// Mitsubishi GX Works2 project: V2   PLC: FX3U/FX3UC

PROGRAM MAIN
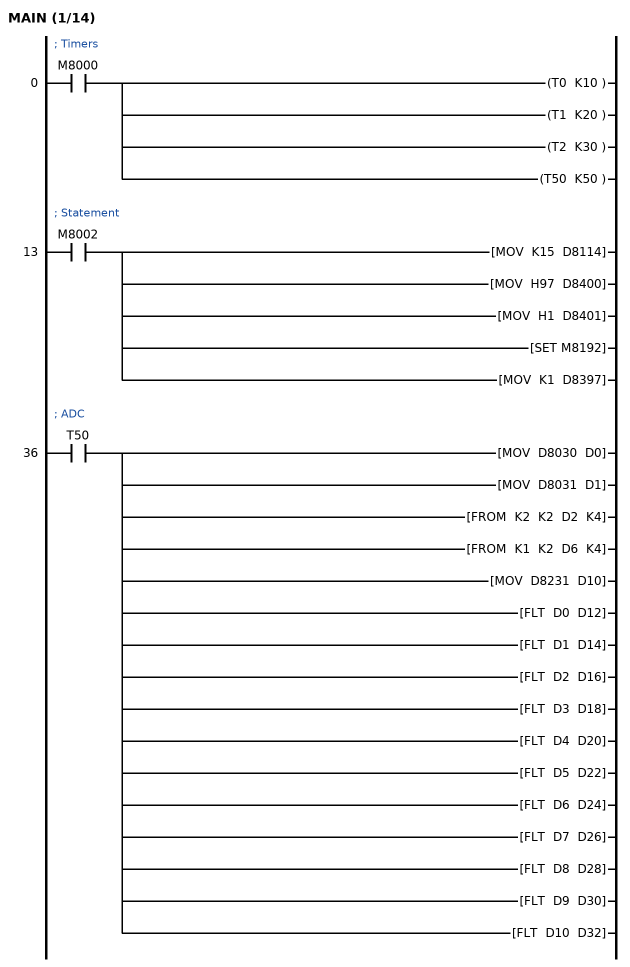
; Timers
0     LD      M8000
      OUT     T0 K10
      OUT     T1 K20
      OUT     T2 K30
      OUT     T50 K50
; Statement
13    LD      M8002
      MOV     K15 D8114
      MOV     H97 D8400
      MOV     H1 D8401
      SET     M8192
      MOV     K1 D8397
; ADC
36    LD      T50
      MOV     D8030 D0
      MOV     D8031 D1
      FROM    K2 K2 D2 K4
      FROM    K1 K2 D6 K4
      MOV     D8231 D10
      FLT     D0 D12
      FLT     D1 D14
      FLT     D2 D16
      FLT     D3 D18
      FLT     D4 D20
      FLT     D5 D22
      FLT     D6 D24
      FLT     D7 D26
      FLT     D8 D28
      FLT     D9 D30
      FLT     D10 D32
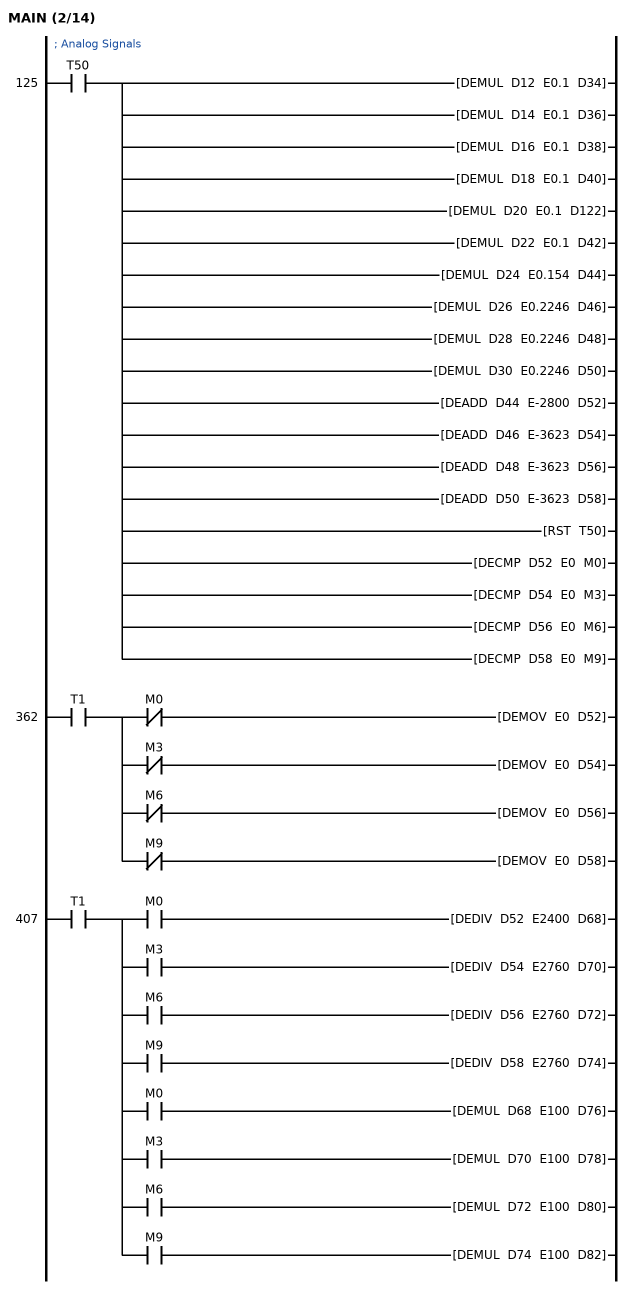
; Analog Signals
125   LD      T50
      DEMUL   D12 E0.1 D34
      DEMUL   D14 E0.1 D36
      DEMUL   D16 E0.1 D38
      DEMUL   D18 E0.1 D40
      DEMUL   D20 E0.1 D122
      DEMUL   D22 E0.1 D42
      DEMUL   D24 E0.154 D44
      DEMUL   D26 E0.2246 D46
      DEMUL   D28 E0.2246 D48
      DEMUL   D30 E0.2246 D50
      DEADD   D44 E-2800 D52
      DEADD   D46 E-3623 D54
      DEADD   D48 E-3623 D56
      DEADD   D50 E-3623 D58
      RST     T50
      DECMP   D52 E0 M0
      DECMP   D54 E0 M3
      DECMP   D56 E0 M6
      DECMP   D58 E0 M9
362   LD      T1
      MPS
      ANI     M0
      DEMOV   E0 D52
      MRD
      ANI     M3
      DEMOV   E0 D54
      MRD
      ANI     M6
      DEMOV   E0 D56
      MPP
      ANI     M9
      DEMOV   E0 D58
407   LD      T1
      MPS
      AND     M0
      DEDIV   D52 E2400 D68
      MRD
      AND     M3
      DEDIV   D54 E2760 D70
      MRD
      AND     M6
      DEDIV   D56 E2760 D72
      MRD
      AND     M9
      DEDIV   D58 E2760 D74
      MRD
      AND     M0
      DEMUL   D68 E100 D76
      MRD
      AND     M3
      DEMUL   D70 E100 D78
      MRD
      AND     M6
      DEMUL   D72 E100 D80
      MPP
      AND     M9
      DEMUL   D74 E100 D82
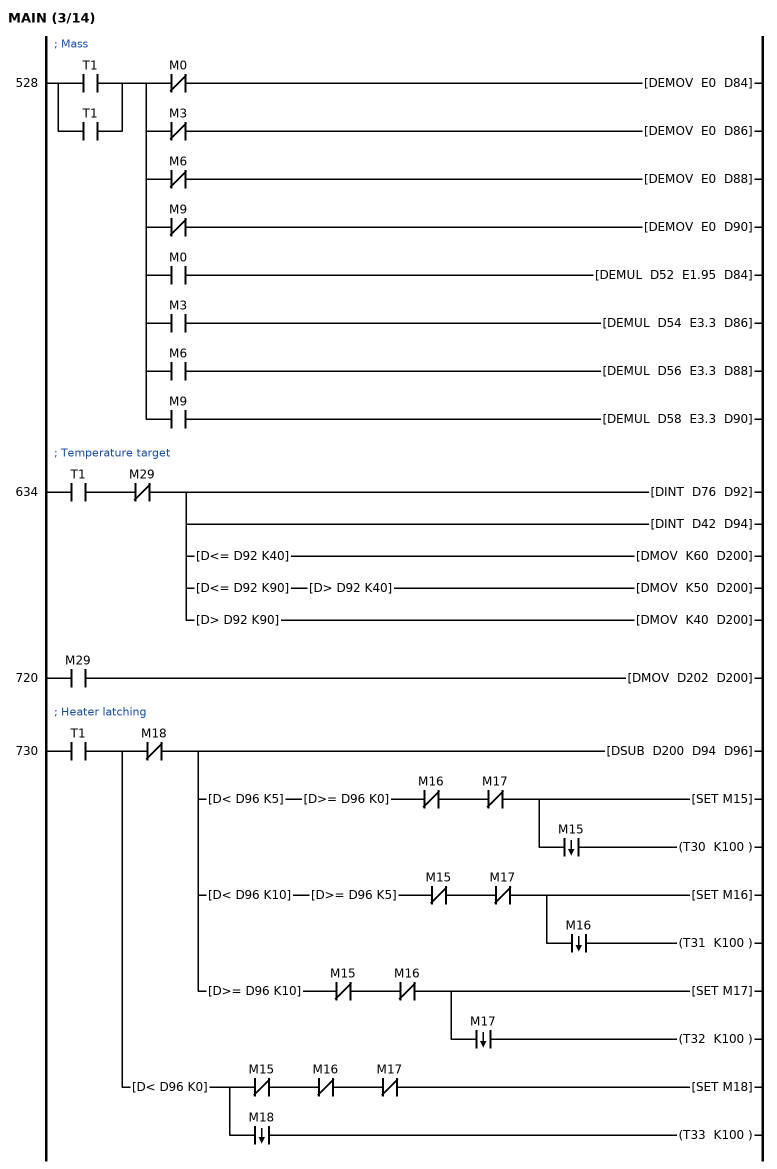
; Mass
528   LD      T1
      OR      T1
      MPS
      ANI     M0
      DEMOV   E0 D84
      MRD
      ANI     M3
      DEMOV   E0 D86
      MRD
      ANI     M6
      DEMOV   E0 D88
      MRD
      ANI     M9
      DEMOV   E0 D90
      MRD
      AND     M0
      DEMUL   D52 E1.95 D84
      MRD
      AND     M3
      DEMUL   D54 E3.3 D86
      MRD
      AND     M6
      DEMUL   D56 E3.3 D88
      MPP
      AND     M9
      DEMUL   D58 E3.3 D90
; Temperature target
634   LD      T1
      ANI     M29
      DINT    D76 D92
      DINT    D42 D94
      MPS
      ANDD<=  D92 K40
      DMOV    K60 D200
      MRD
      ANDD<=  D92 K90
      ANDD>   D92 K40
      DMOV    K50 D200
      MPP
      ANDD>   D92 K90
      DMOV    K40 D200
720   LD      M29
      DMOV    D202 D200
; Heater latching
730   LD      T1
      MPS
      ANI     M18
      DSUB    D200 D94 D96
      MPS
      ANDD<   D96 K5
      ANDD>=  D96 K0
      ANI     M16
      ANI     M17
      SET     M15
      ANDF    M15
      OUT     T30 K100
      MRD
      ANDD<   D96 K10
      ANDD>=  D96 K5
      ANI     M15
      ANI     M17
      SET     M16
      ANDF    M16
      OUT     T31 K100
      MPP
      ANDD>=  D96 K10
      ANI     M15
      ANI     M16
      SET     M17
      ANDF    M17
      OUT     T32 K100
      MPP
      ANDD<   D96 K0
      MPS
      ANI     M15
      ANI     M16
      ANI     M17
      SET     M18
      MPP
      ANDF    M18
      OUT     T33 K100
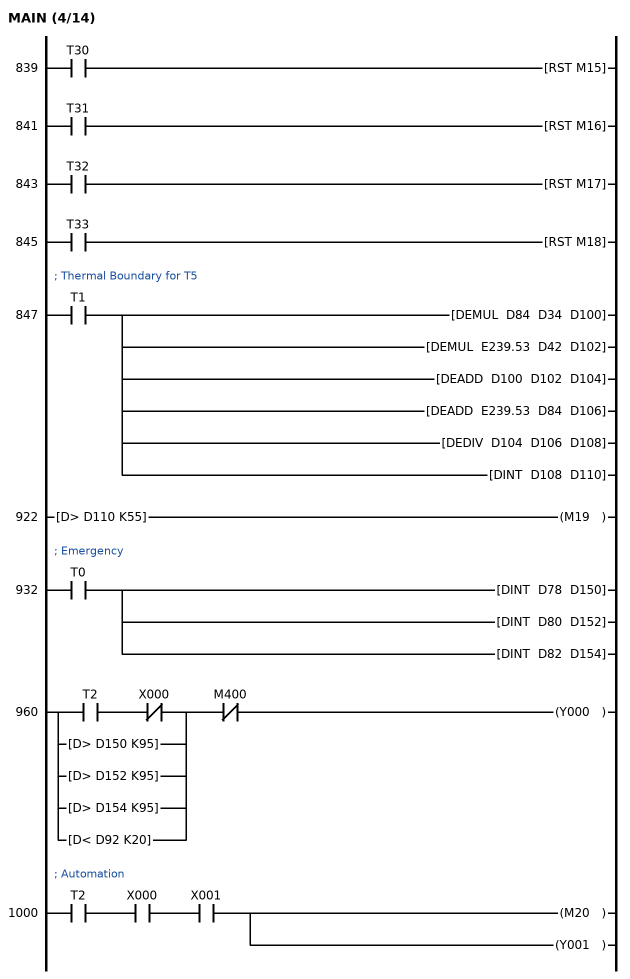
839   LD      T30
      RST     M15
841   LD      T31
      RST     M16
843   LD      T32
      RST     M17
845   LD      T33
      RST     M18
; Thermal Boundary for T5
847   LD      T1
      DEMUL   D84 D34 D100
      DEMUL   E239.53 D42 D102
      DEADD   D100 D102 D104
      DEADD   E239.53 D84 D106
      DEDIV   D104 D106 D108
      DINT    D108 D110
922   LDD>    D110 K55
      OUT     M19
; Emergency
932   LD      T0
      DINT    D78 D150
      DINT    D80 D152
      DINT    D82 D154
960   LD      T2
      ANI     X000
      ORD>    D150 K95
      ORD>    D152 K95
      ORD>    D154 K95
      ORD<    D92 K20
      ANI     M400
      OUT     Y000
; Automation
1000  LD      T2
      AND     X000
      AND     X001
      OUT     M20
      OUT     Y001
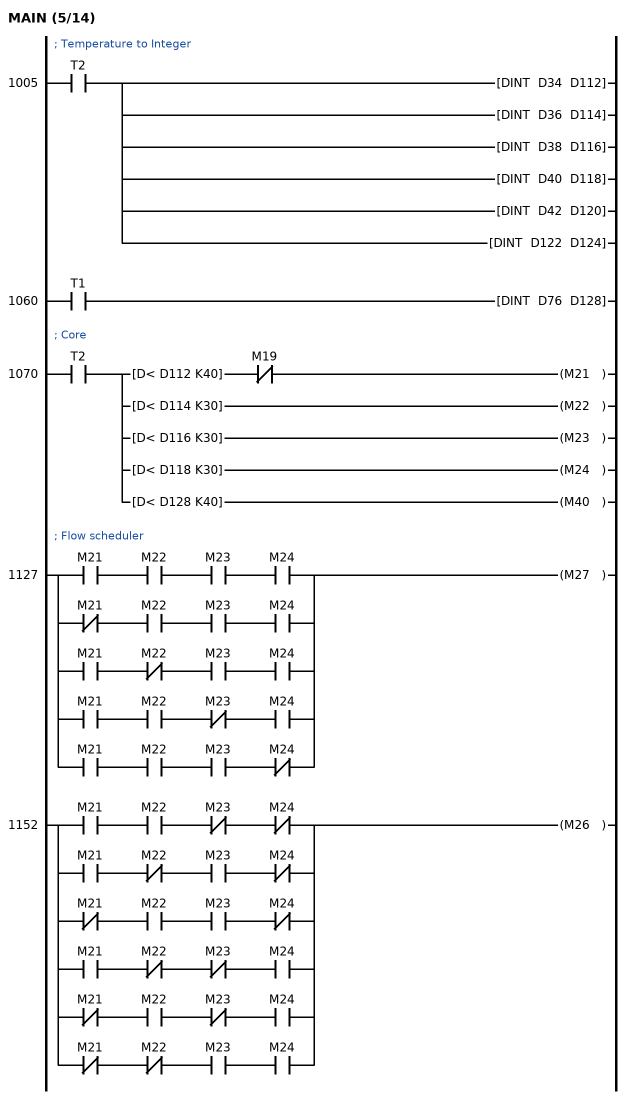
; Temperature to Integer
1005  LD      T2
      DINT    D34 D112
      DINT    D36 D114
      DINT    D38 D116
      DINT    D40 D118
      DINT    D42 D120
      DINT    D122 D124
1060  LD      T1
      DINT    D76 D128
; Core
1070  LD      T2
      MPS
      ANDD<   D112 K40
      ANI     M19
      OUT     M21
      MRD
      ANDD<   D114 K30
      OUT     M22
      MRD
      ANDD<   D116 K30
      OUT     M23
      MRD
      ANDD<   D118 K30
      OUT     M24
      MPP
      ANDD<   D128 K40
      OUT     M40
; Flow scheduler
1127  LD      M21
      AND     M22
      AND     M23
      AND     M24
      LDI     M21
      AND     M22
      AND     M23
      AND     M24
      ORB
      LD      M21
      ANI     M22
      AND     M23
      AND     M24
      ORB
      LD      M21
      AND     M22
      ANI     M23
      AND     M24
      ORB
      LD      M21
      AND     M22
      AND     M23
      ANI     M24
      ORB
      OUT     M27
1152  LD      M21
      AND     M22
      ANI     M23
      ANI     M24
      LD      M21
      ANI     M22
      AND     M23
      ANI     M24
      ORB
      LDI     M21
      AND     M22
      AND     M23
      ANI     M24
      ORB
      LD      M21
      ANI     M22
      ANI     M23
      AND     M24
      ORB
      LDI     M21
      AND     M22
      ANI     M23
      AND     M24
      ORB
      LDI     M21
      ANI     M22
      AND     M23
      AND     M24
      ORB
      OUT     M26
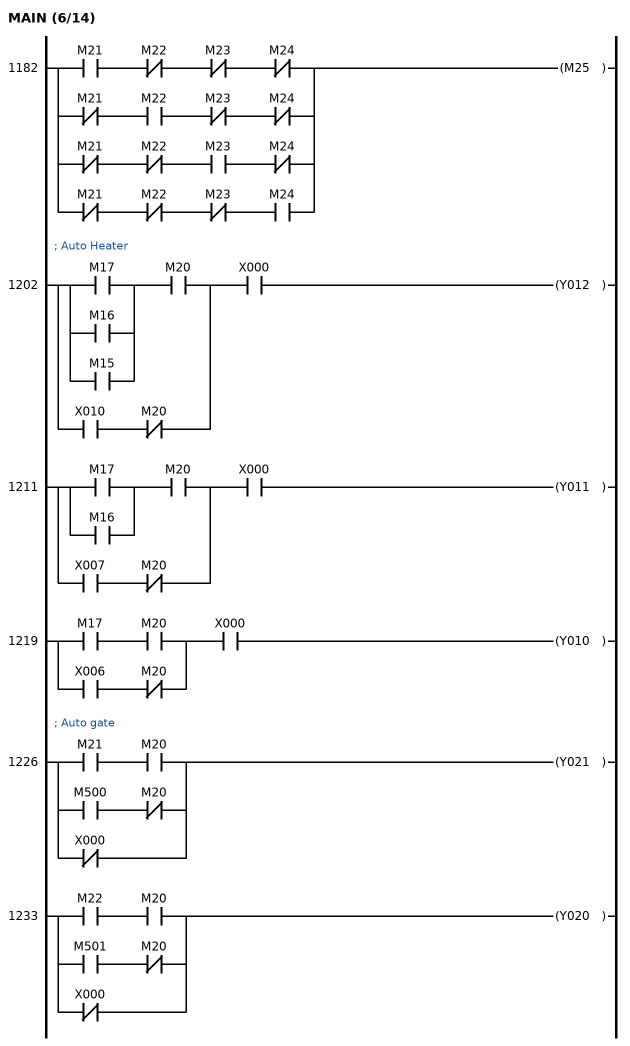
1182  LD      M21
      ANI     M22
      ANI     M23
      ANI     M24
      LDI     M21
      AND     M22
      ANI     M23
      ANI     M24
      ORB
      LDI     M21
      ANI     M22
      AND     M23
      ANI     M24
      ORB
      LDI     M21
      ANI     M22
      ANI     M23
      AND     M24
      ORB
      OUT     M25
; Auto Heater
1202  LD      M17
      OR      M16
      OR      M15
      AND     M20
      LD      X010
      ANI     M20
      ORB
      AND     X000
      OUT     Y012
1211  LD      M17
      OR      M16
      AND     M20
      LD      X007
      ANI     M20
      ORB
      AND     X000
      OUT     Y011
1219  LD      M17
      AND     M20
      LD      X006
      ANI     M20
      ORB
      AND     X000
      OUT     Y010
; Auto gate
1226  LD      M21
      AND     M20
      LD      M500
      ANI     M20
      ORB
      ORI     X000
      OUT     Y021
1233  LD      M22
      AND     M20
      LD      M501
      ANI     M20
      ORB
      ORI     X000
      OUT     Y020
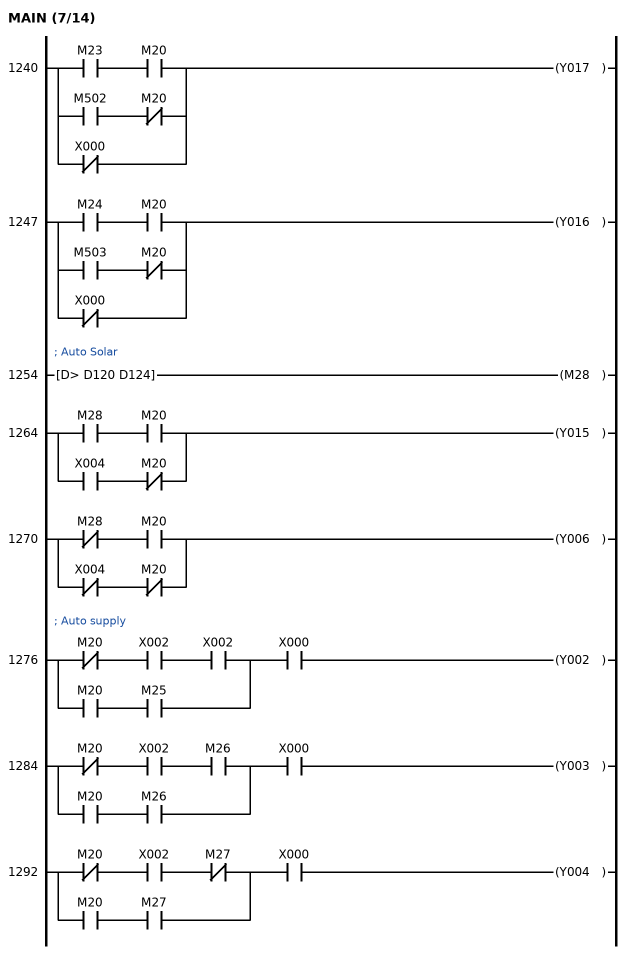
1240  LD      M23
      AND     M20
      LD      M502
      ANI     M20
      ORB
      ORI     X000
      OUT     Y017
1247  LD      M24
      AND     M20
      LD      M503
      ANI     M20
      ORB
      ORI     X000
      OUT     Y016
; Auto Solar
1254  LDD>    D120 D124
      OUT     M28
1264  LD      M28
      AND     M20
      LD      X004
      ANI     M20
      ORB
      OUT     Y015
1270  LDI     M28
      AND     M20
      LDI     X004
      ANI     M20
      ORB
      OUT     Y006
; Auto supply
1276  LDI     M20
      AND     X002
      AND     X002
      LD      M20
      AND     M25
      ORB
      AND     X000
      OUT     Y002
1284  LDI     M20
      AND     X002
      AND     M26
      LD      M20
      AND     M26
      ORB
      AND     X000
      OUT     Y003
1292  LDI     M20
      AND     X002
      ANI     M27
      LD      M20
      AND     M27
      ORB
      AND     X000
      OUT     Y004
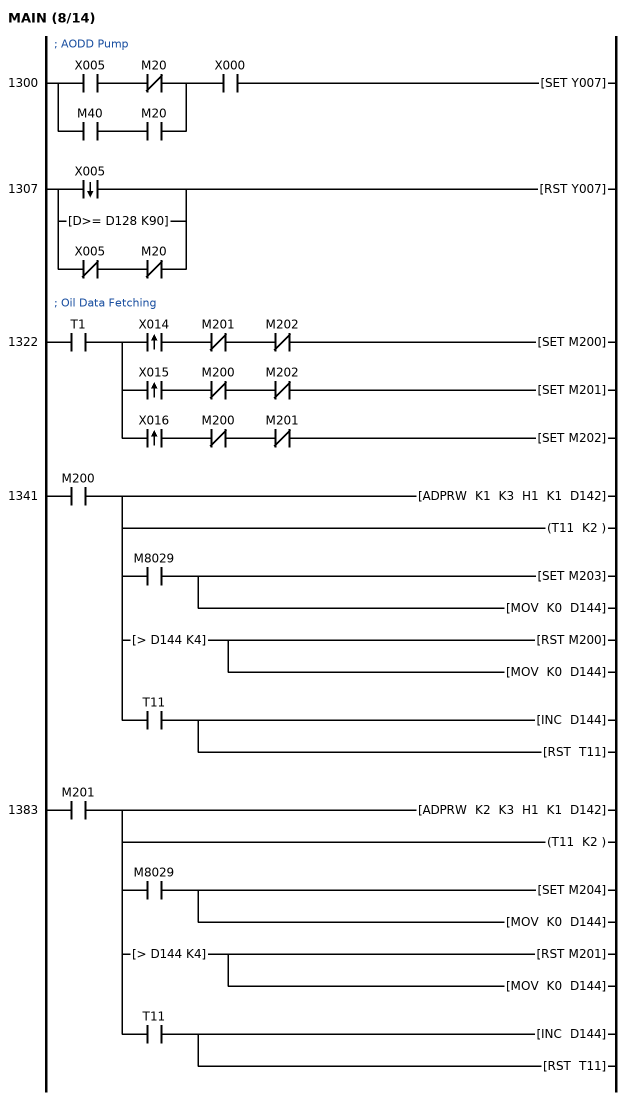
; AODD Pump
1300  LD      X005
      ANI     M20
      LD      M40
      AND     M20
      ORB
      AND     X000
      SET     Y007
1307  LDF     X005
      ORD>=   D128 K90
      LDI     X005
      ANI     M20
      ORB
      RST     Y007
; Oil Data Fetching
1322  LD      T1
      MPS
      ANDP    X014
      ANI     M201
      ANI     M202
      SET     M200
      MRD
      ANDP    X015
      ANI     M200
      ANI     M202
      SET     M201
      MPP
      ANDP    X016
      ANI     M200
      ANI     M201
      SET     M202
1341  LD      M200
      ADPRW   K1 K3 H1 K1 D142
      OUT     T11 K2
      MPS
      AND     M8029
      SET     M203
      MOV     K0 D144
      MRD
      AND>    D144 K4
      RST     M200
      MOV     K0 D144
      MPP
      AND     T11
      INC     D144
      RST     T11
1383  LD      M201
      ADPRW   K2 K3 H1 K1 D142
      OUT     T11 K2
      MPS
      AND     M8029
      SET     M204
      MOV     K0 D144
      MRD
      AND>    D144 K4
      RST     M201
      MOV     K0 D144
      MPP
      AND     T11
      INC     D144
      RST     T11
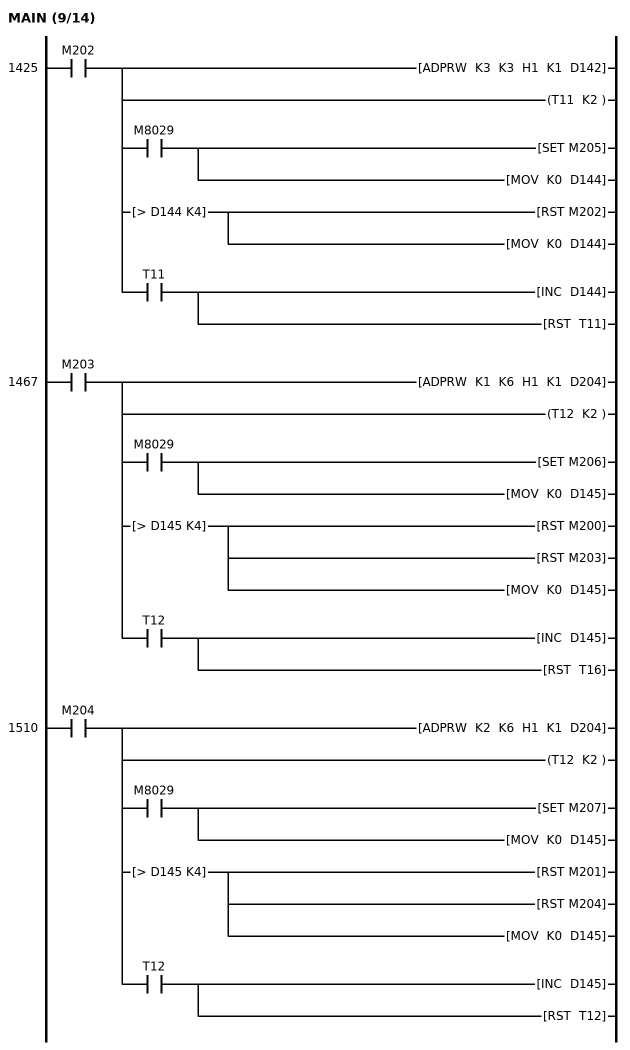
1425  LD      M202
      ADPRW   K3 K3 H1 K1 D142
      OUT     T11 K2
      MPS
      AND     M8029
      SET     M205
      MOV     K0 D144
      MRD
      AND>    D144 K4
      RST     M202
      MOV     K0 D144
      MPP
      AND     T11
      INC     D144
      RST     T11
1467  LD      M203
      ADPRW   K1 K6 H1 K1 D204
      OUT     T12 K2
      MPS
      AND     M8029
      SET     M206
      MOV     K0 D145
      MRD
      AND>    D145 K4
      RST     M200
      RST     M203
      MOV     K0 D145
      MPP
      AND     T12
      INC     D145
      RST     T16
1510  LD      M204
      ADPRW   K2 K6 H1 K1 D204
      OUT     T12 K2
      MPS
      AND     M8029
      SET     M207
      MOV     K0 D145
      MRD
      AND>    D145 K4
      RST     M201
      RST     M204
      MOV     K0 D145
      MPP
      AND     T12
      INC     D145
      RST     T12
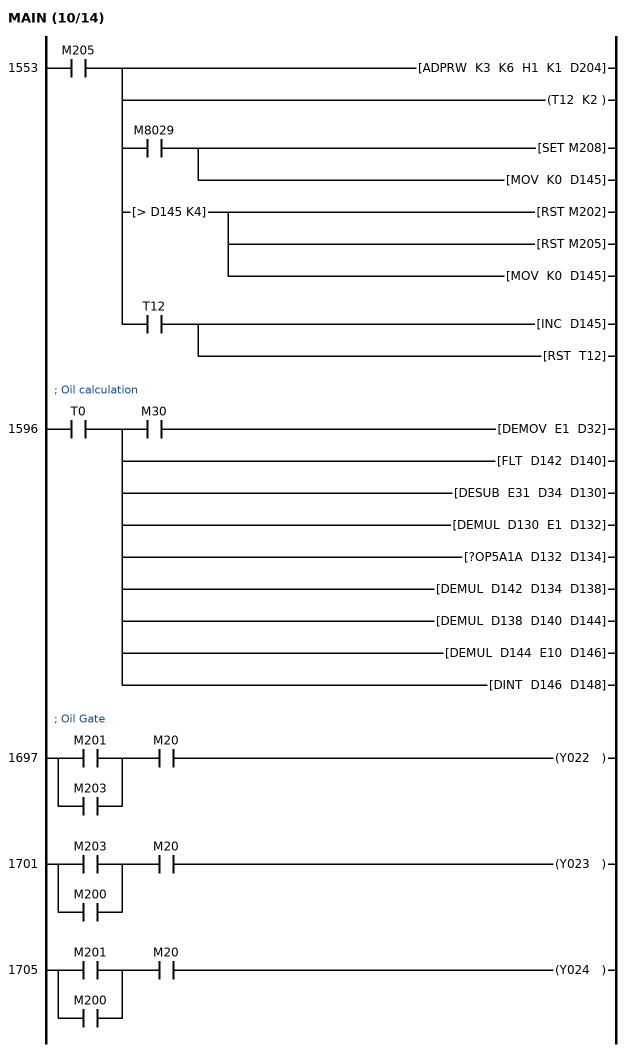
1553  LD      M205
      ADPRW   K3 K6 H1 K1 D204
      OUT     T12 K2
      MPS
      AND     M8029
      SET     M208
      MOV     K0 D145
      MRD
      AND>    D145 K4
      RST     M202
      RST     M205
      MOV     K0 D145
      MPP
      AND     T12
      INC     D145
      RST     T12
; Oil calculation
1596  LD      T0
      MPS
      AND     M30
      DEMOV   E1 D32
      MPP
      FLT     D142 D140
      DESUB   E31 D34 D130
      DEMUL   D130 E1 D132
      ?OP5A1A D132 D134
      DEMUL   D142 D134 D138
      DEMUL   D138 D140 D144
      DEMUL   D144 E10 D146
      DINT    D146 D148
; Oil Gate
1697  LD      M201
      OR      M203
      AND     M20
      OUT     Y022
1701  LD      M203
      OR      M200
      AND     M20
      OUT     Y023
1705  LD      M201
      OR      M200
      AND     M20
      OUT     Y024
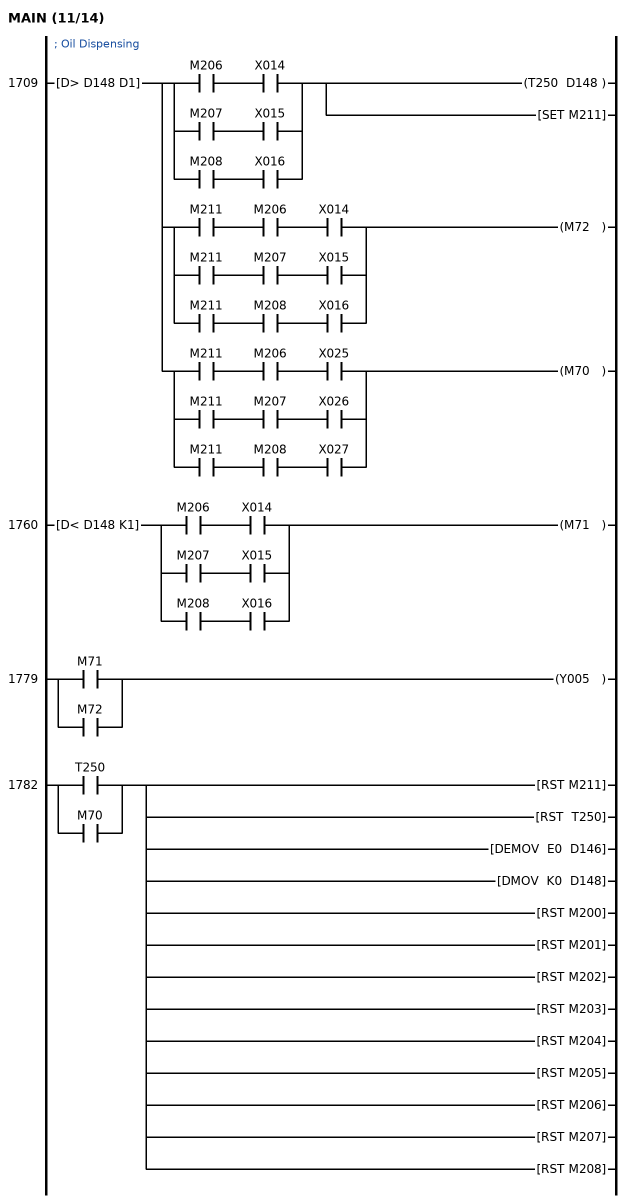
; Oil Dispensing
1709  LDD>    D148 D1
      MPS
      LD      M206
      AND     X014
      LD      M207
      AND     X015
      ORB
      LD      M208
      AND     X016
      ORB
      ANB
      OUT     T250 D148
      SET     M211
      MRD
      LD      M211
      AND     M206
      AND     X014
      LD      M211
      AND     M207
      AND     X015
      ORB
      LD      M211
      AND     M208
      AND     X016
      ORB
      ANB
      OUT     M72
      MPP
      LD      M211
      AND     M206
      AND     X025
      LD      M211
      AND     M207
      AND     X026
      ORB
      LD      M211
      AND     M208
      AND     X027
      ORB
      ANB
      OUT     M70
1760  LDD<    D148 K1
      LD      M206
      AND     X014
      LD      M207
      AND     X015
      ORB
      LD      M208
      AND     X016
      ORB
      ANB
      OUT     M71
1779  LD      M71
      OR      M72
      OUT     Y005
1782  LD      T250
      OR      M70
      RST     M211
      RST     T250
      DEMOV   E0 D146
      DMOV    K0 D148
      RST     M200
      RST     M201
      RST     M202
      RST     M203
      RST     M204
      RST     M205
      RST     M206
      RST     M207
      RST     M208
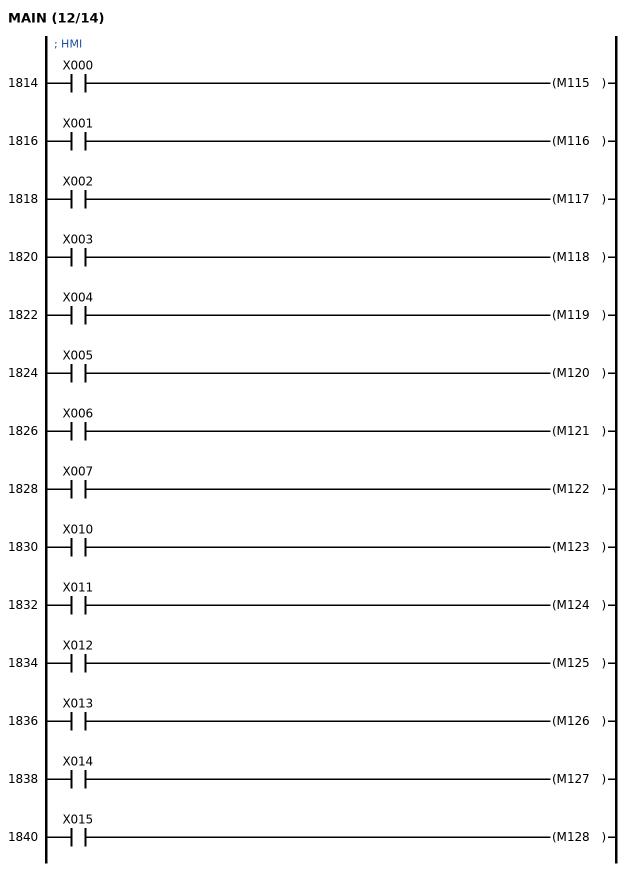
; HMI
1814  LD      X000
      OUT     M115
1816  LD      X001
      OUT     M116
1818  LD      X002
      OUT     M117
1820  LD      X003
      OUT     M118
1822  LD      X004
      OUT     M119
1824  LD      X005
      OUT     M120
1826  LD      X006
      OUT     M121
1828  LD      X007
      OUT     M122
1830  LD      X010
      OUT     M123
1832  LD      X011
      OUT     M124
1834  LD      X012
      OUT     M125
1836  LD      X013
      OUT     M126
1838  LD      X014
      OUT     M127
1840  LD      X015
      OUT     M128
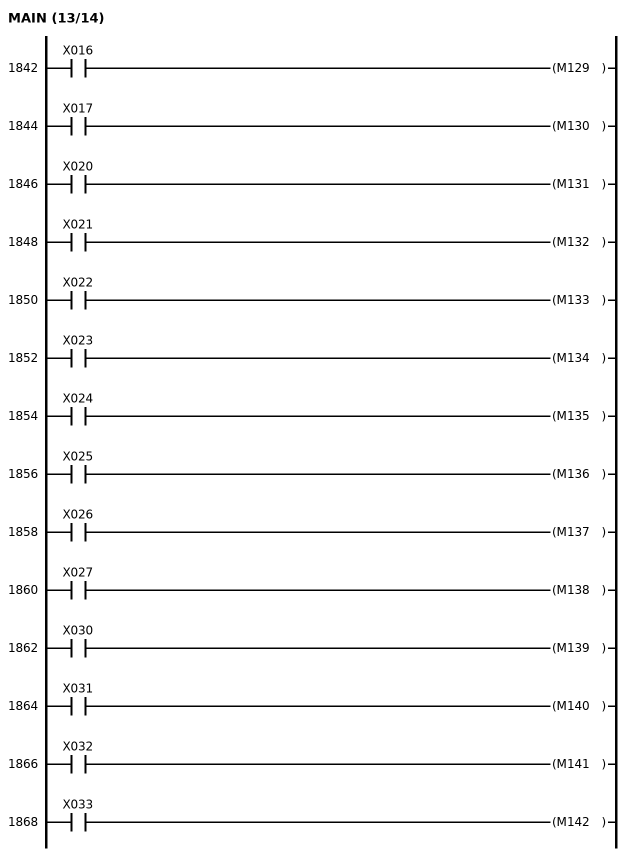
1842  LD      X016
      OUT     M129
1844  LD      X017
      OUT     M130
1846  LD      X020
      OUT     M131
1848  LD      X021
      OUT     M132
1850  LD      X022
      OUT     M133
1852  LD      X023
      OUT     M134
1854  LD      X024
      OUT     M135
1856  LD      X025
      OUT     M136
1858  LD      X026
      OUT     M137
1860  LD      X027
      OUT     M138
1862  LD      X030
      OUT     M139
1864  LD      X031
      OUT     M140
1866  LD      X032
      OUT     M141
1868  LD      X033
      OUT     M142
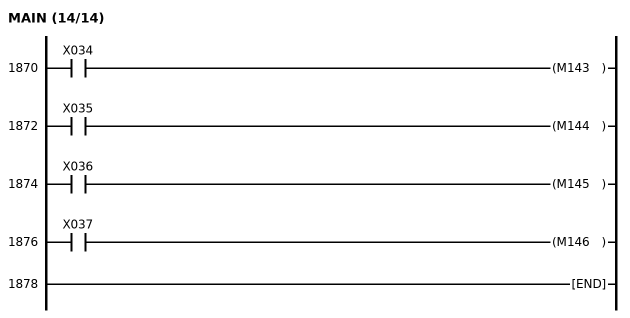
1870  LD      X034
      OUT     M143
1872  LD      X035
      OUT     M144
1874  LD      X036
      OUT     M145
1876  LD      X037
      OUT     M146
1878  END
END_PROGRAM
